FUNCTION_BLOCK VALVE_FEEDBACK (* Migrated from IEC 61131-3 ST *)
  (* Standard: 61499-2 *)
  (* Version 1.0, 2026-11-06, st2fb *)
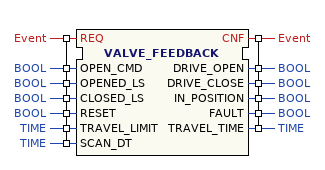
  EVENT_INPUT
    REQ WITH OPEN_CMD, OPENED_LS, CLOSED_LS, RESET, TRAVEL_LIMIT, SCAN_DT;
  END_EVENT
  EVENT_OUTPUT
    CNF WITH DRIVE_OPEN, DRIVE_CLOSE, IN_POSITION, FAULT, TRAVEL_TIME;
  END_EVENT
  VAR_INPUT
    OPEN_CMD : BOOL;
    OPENED_LS : BOOL;
    CLOSED_LS : BOOL;
    RESET : BOOL;
    TRAVEL_LIMIT : TIME;
    SCAN_DT : TIME;
  END_VAR
  VAR_OUTPUT
    DRIVE_OPEN : BOOL;
    DRIVE_CLOSE : BOOL;
    IN_POSITION : BOOL;
    FAULT : BOOL;
    TRAVEL_TIME : TIME;
  END_VAR
  VAR
    ST2FB_NOW : TIME := T#0s;
    OPENING_TIMER_IN : BOOL;
    OPENING_TIMER_PT : TIME;
    OPENING_TIMER_Q : BOOL;
    OPENING_TIMER_ET : TIME;
    OPENING_TIMER_STATE : INT;
    OPENING_TIMER_PREV_IN : BOOL;
    OPENING_TIMER_START_TIME : TIME;
    CLOSING_TIMER_IN : BOOL;
    CLOSING_TIMER_PT : TIME;
    CLOSING_TIMER_Q : BOOL;
    CLOSING_TIMER_ET : TIME;
    CLOSING_TIMER_STATE : INT;
    CLOSING_TIMER_PREV_IN : BOOL;
    CLOSING_TIMER_START_TIME : TIME;
  END_VAR
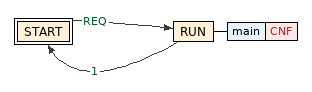
  EC_STATES
    START;
    RUN : main -> CNF;
  END_STATES
  EC_TRANSITIONS
    START TO RUN := REQ;
    RUN TO START := 1;
  END_TRANSITIONS
  ALGORITHM main IN ST:
ST2FB_NOW := ST2FB_NOW + SCAN_DT;

OPENING_TIMER_IN := OPEN_CMD AND NOT OPENED_LS;
OPENING_TIMER_PT := TRAVEL_LIMIT;
IF (OPENING_TIMER_STATE = 0) AND NOT OPENING_TIMER_PREV_IN AND OPENING_TIMER_IN THEN
  OPENING_TIMER_STATE := 1;
  OPENING_TIMER_Q := FALSE;
  OPENING_TIMER_START_TIME := ST2FB_NOW;
ELSE
  IF NOT OPENING_TIMER_IN THEN
    OPENING_TIMER_ET := T#0s;
    OPENING_TIMER_Q := FALSE;
    OPENING_TIMER_STATE := 0;
  ELSIF OPENING_TIMER_STATE = 1 THEN
    IF OPENING_TIMER_START_TIME + OPENING_TIMER_PT <= ST2FB_NOW THEN
      OPENING_TIMER_STATE := 2;
      OPENING_TIMER_Q := TRUE;
      OPENING_TIMER_ET := OPENING_TIMER_PT;
    ELSE
      OPENING_TIMER_ET := ST2FB_NOW - OPENING_TIMER_START_TIME;
    END_IF;
  END_IF;
END_IF;
OPENING_TIMER_PREV_IN := OPENING_TIMER_IN;

CLOSING_TIMER_IN := NOT OPEN_CMD AND NOT CLOSED_LS;
CLOSING_TIMER_PT := TRAVEL_LIMIT;
IF (CLOSING_TIMER_STATE = 0) AND NOT CLOSING_TIMER_PREV_IN AND CLOSING_TIMER_IN THEN
  CLOSING_TIMER_STATE := 1;
  CLOSING_TIMER_Q := FALSE;
  CLOSING_TIMER_START_TIME := ST2FB_NOW;
ELSE
  IF NOT CLOSING_TIMER_IN THEN
    CLOSING_TIMER_ET := T#0s;
    CLOSING_TIMER_Q := FALSE;
    CLOSING_TIMER_STATE := 0;
  ELSIF CLOSING_TIMER_STATE = 1 THEN
    IF CLOSING_TIMER_START_TIME + CLOSING_TIMER_PT <= ST2FB_NOW THEN
      CLOSING_TIMER_STATE := 2;
      CLOSING_TIMER_Q := TRUE;
      CLOSING_TIMER_ET := CLOSING_TIMER_PT;
    ELSE
      CLOSING_TIMER_ET := ST2FB_NOW - CLOSING_TIMER_START_TIME;
    END_IF;
  END_IF;
END_IF;
CLOSING_TIMER_PREV_IN := CLOSING_TIMER_IN;

IF OPENING_TIMER_Q OR CLOSING_TIMER_Q OR (OPENED_LS AND CLOSED_LS) THEN
  FAULT := TRUE;
ELSIF RESET THEN
  FAULT := FALSE;
END_IF;
DRIVE_OPEN := OPEN_CMD AND NOT OPENED_LS AND NOT FAULT;
DRIVE_CLOSE := NOT OPEN_CMD AND NOT CLOSED_LS AND NOT FAULT;
IN_POSITION := NOT FAULT AND ((OPEN_CMD AND OPENED_LS) OR (NOT OPEN_CMD AND CLOSED_LS));
IF OPEN_CMD THEN
  TRAVEL_TIME := OPENING_TIMER_ET;
ELSE
  TRAVEL_TIME := CLOSING_TIMER_ET;
END_IF;
  END_ALGORITHM
END_FUNCTION_BLOCK
